PROGRAM Zabezpieczenie_Tensometru
VAR
	bPrzeciazenieTensometru: BOOL;
	rtOverload: R_TRIG;
END_VAR

IF GVL_ForceMode.bForceRange100t=0 THEN
	IF GVL_ForceMode.nForce_t>51 THEN 
		bPrzeciazenieTensometru:=TRUE;
	END_IF
END_IF
IF GVL_ForceMode.bForceRange100t=1 THEN
	IF GVL_ForceMode.nForce_t>101 THEN 
		bPrzeciazenieTensometru:=TRUE;
	END_IF
END_IF

rtOverload(CLK:=bPrzeciazenieTensometru , Q=> );

END_PROGRAM

(* stored: Version 1.1.0.1, ProductVersion 3.1.4024.16
   POU Zabezpieczenie_Tensometru: Id {b9123738-7943-47bb-8681-d725bfd74512}, SpecialFunc None *)
